Fanuc KAREL source: kd00030.KL

-- PROVISIONAL review KL for V770-1; original PC SHA256 59c98dabb68fbd149f2cab6097680936436a8164ee854c3c34f6642dd08d6be8
-- Incomplete behavior may be omitted. Consult companion uncertainty JSON. Do not deploy.
PROGRAM KD00030
%NOLOCKGROUP
VAR
  I : INTEGER
  J : INTEGER
  B : BOOLEAN
  R : REAL
  S : STRING[80]
BEGIN
  -- UNRESOLVED_PC offsets 5-21; opcodes 9D,81,18,9C,12,22,9D,13,04
  -- UNRESOLVED_PC offsets 26-30; opcodes 7F
END KD00030
